Staubli VAL3: load.pgx

program load()
  local string l_sPath
  local bool l_bResult
  local num l_nResult
begin
//call trajectory:loadTRAJ(savedata:nLibIndex,l_nResult)
end
